KUKA KRL data list: folge11.dat

&ACCESS RVP
&REL 1
&COMMENT bt2krl sim data Folge 11 plan 16#A312
DEFDAT FOLGE11
   ; Generated by bt2krl 0.1.0 from bt2plc plan bt_1791274820_cell_2robot (cell cell_2robot), PLAN_ID 16#A312
   ; Robot robot1 (R1), controller robot1, model KR240R2900_ULTRA, joint mapping identity
   ; Profile sim (bt2plc simulator telegram). NEVER install on a VW KS24 robot:
   ; its signals collide with the VW standard (Fertigmeldung, interlocks, PRG_NR).
   ; Do not edit: regenerate with bt2krl (plain KRL, no inline forms).
   EXT BAS (BAS_COMMAND :IN,REAL :IN )
   DECL INT PLAN_ID=41746
   DECL AXIS P1={A1 0.0,A2 -90.0,A3 90.0,A4 0.0,A5 0.0,A6 0.0}
   DECL AXIS P2={A1 0.1421,A2 -89.0006,A3 89.9771,A4 0.0,A5 0.0,A6 0.0}
   DECL AXIS P3={A1 0.5354,A2 -86.231,A3 89.9133,A4 0.0,A5 0.0,A6 0.0}
   DECL AXIS P4={A1 1.131,A2 -82.0342,A3 89.8161,A4 0.0,A5 0.0,A6 0.0}
   DECL AXIS P5={A1 1.8795,A2 -76.7531,A3 89.6931,A4 0.0,A5 0.0,A6 0.0}
   DECL AXIS P6={A1 5.42,A2 -51.6436,A3 89.0908,A4 0.0,A5 0.0,A6 0.0}
   DECL AXIS P7={A1 6.1959,A2 -46.0847,A3 88.9501,A4 0.0,A5 0.0,A6 0.0}
   DECL AXIS P8={A1 6.8297,A2 -41.499,A3 88.8283,A4 0.0,A5 0.0,A6 0.0}
   DECL AXIS P9={A1 7.2722,A2 -38.2294,A3 88.7329,A4 0.0,A5 0.0,A6 0.0}
   DECL AXIS P10={A1 7.7267,A2 -33.2119,A3 88.3788,A4 0.0,A5 0.0,A6 0.0}
   DECL AXIS P11={A1 7.2722,A2 -35.0616,A3 88.2443,A4 0.0,A5 0.0,A6 0.0}
   DECL AXIS P12={A1 7.1292,A2 -36.1426,A3 88.2788,A4 0.0,A5 0.0,A6 0.0}
   DECL AXIS P13={A1 6.7336,A2 -39.1311,A3 88.3743,A4 0.0,A5 0.0,A6 0.0}
   DECL AXIS P14={A1 6.136,A2 -43.6457,A3 88.5186,A4 0.0,A5 0.0,A6 0.0}
   DECL AXIS P15={A1 5.3868,A2 -49.3049,A3 88.6995,A4 0.0,A5 0.0,A6 0.0}
   DECL AXIS P16={A1 1.8854,A2 -75.7567,A3 89.5448,A4 0.0,A5 0.0,A6 0.0}
   DECL AXIS P17={A1 1.1363,A2 -81.4159,A3 89.7257,A4 0.0,A5 0.0,A6 0.0}
   DECL AXIS P18={A1 0.5387,A2 -85.9305,A3 89.8699,A4 0.0,A5 0.0,A6 0.0}
   DECL AXIS P19={A1 0.1431,A2 -88.919,A3 89.9655,A4 0.0,A5 0.0,A6 0.0}
   DECL AXIS P20={A1 0.0,A2 -90.0,A3 90.0,A4 0.0,A5 0.0,A6 0.0}
ENDDAT
